// TIA Portal V19 export
// export: Created 2026-11-24T14:48:46.8883601Z, ExportSetting WithDefaults, DisplayName Totally Integrated Automation Portal, DisplayVersion V19, DisplayName TIA Portal Openness, DisplayVersion V19, DisplayName TIA Portal Version Control Interface, DisplayVersion V19, DisplayName STEP 7 Professional, DisplayVersion V19, DisplayName STEP 7 Safety, DisplayVersion V19, DisplayName WinCC Basic/Comfort/Advanced, DisplayVersion V19, DisplayName WinCC Unified, DisplayVersion V19
VAR_GLOBAL   // PLC tag table "Farm_IO"
   DI_EStopOk AT %I0.0 : Bool;   // E-stop circuit healthy (NC; FALSE = pressed)
   DI_MainsOk AT %I0.1 : Bool;   // Mains present (relay before the UPS)
   DI_BoosterRun AT %I0.2 : Bool;   // Booster running
   DI_BoosterFault AT %I0.3 : Bool;   // Booster overload / drive fault
   DI_WellRun AT %I0.4 : Bool;   // Well pump running
   DI_WellFault AT %I0.5 : Bool;   // Well pump overload / drive fault
   DI_BoosterHand AT %I0.6 : Bool;   // Booster selector HAND
   DI_BoosterOff AT %I0.7 : Bool;   // Booster selector OFF
   DI_WellHand AT %I1.0 : Bool;   // Well selector HAND
   DI_WellOff AT %I1.1 : Bool;   // Well selector OFF
   DI_ZoneOnLo AT %IB2 : Byte;   // Zone selectors 1-8 ON
   DI_ZoneOnHi AT %IB3 : Byte;   // Zone selectors 9-16 ON
   DI_ZoneOffLo AT %IB4 : Byte;   // Zone selectors 1-8 OFF
   DI_ZoneOffHi AT %IB5 : Byte;   // Zone selectors 9-16 OFF
   AI_TankLevel AT %IW6 : Int;   // Tank level 4-20 mA
   AI_MainPressure AT %IW8 : Int;   // Mainline pressure 4-20 mA
   AI_MainFlow AT %IW10 : Int;   // Mainline flow 4-20 mA
   AI_WellLevel AT %IW12 : Int;   // Well level 4-20 mA
   AI_FilterDp AT %IW14 : Int;   // Filter pressure drop 4-20 mA
   DQ_ValveLo AT %QB0 : Byte;   // Wired zone valves 1-8
   DQ_ValveHi AT %QB1 : Byte;   // Wired zone valves 9-16
   DQ_BoosterStart AT %Q2.0 : Bool;   // Booster start
   DQ_WellStart AT %Q2.1 : Bool;   // Well pump start
   DQ_Beacon AT %Q2.2 : Bool;   // Red alarm beacon
   DQ_Horn AT %Q2.3 : Bool;   // Horn
END_VAR
